Fanuc KAREL source: KD00036.KL

PROGRAM KD00036
%NOLOCKGROUP
VAR
  I: INTEGER
  J: INTEGER
  B: BOOLEAN
  R: REAL
  S: STRING[80]
BEGIN
  CONDITION[1]:
  WHEN DIN[1] = ON DO
    NOMESSAGE
  ENDCONDITION
END KD00036
